ABB RAPID module: Wobj_WO_PasReal.mod

MODULE Wobj_WO_PasReal
	! Points are read in order of declaration.
  ! Please do not change the order of points!

  LOCAL PERS robtarget pWobj_U_PointX1:=[[473.2875,1.359913,422.1007],[0.137335553765297,0.00816564448177814,0.990426778793335,-0.0112673677504063],[0,-1,0,0],[9E+09,9E+09,9E+09,9E+09,9E+09,9E+09]];
	LOCAL PERS robtarget pWobj_U_PointX2:=[[471.808,-132.749,420.8833],[0.137332648038864,0.0081624761223793,0.990427255630493,-0.0112657556310296],[-1,0,-1,0],[9E+09,9E+09,9E+09,9E+09,9E+09,9E+09]];
	LOCAL PERS robtarget pWobj_U_PointY1:=[[335.0285,2.047842,419.1656],[0.137334257364273,0.00816600117832422,0.990426957607269,-0.0112643809989095],[0,-1,0,0],[9E+09,9E+09,9E+09,9E+09,9E+09,9E+09]];

ENDMODULE
